FUNCTION_BLOCK StopPointLogic (* Basic Function Block Type *)
  (* Standard: 61499-2 *)
  (* Version 0.0, 11/22/2026, Schneider Electric, First version *)
  PACKAGE Main;
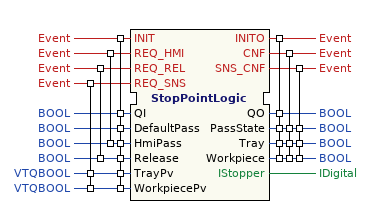
  EVENT_INPUT
    INIT WITH QI, DefaultPass, HmiPass, Release, TrayPv, WorkpiecePv; (* Initialization Request *)
    REQ_HMI WITH HmiPass; (* Update pass-through command from HMI SetBool *)
    REQ_REL WITH Release; (* Update external release request *)
    REQ_SNS WITH TrayPv, WorkpiecePv; (* Update tray and workpiece sensor values *)
  END_EVENT
  EVENT_OUTPUT
    INITO WITH QO, PassState, Tray, Workpiece; (* Initialization Confirm *)
    CNF WITH PassState, Tray, Workpiece; (* Pass-through state confirmation *)
    SNS_CNF WITH Tray, Workpiece, PassState; (* Sensor confirmation *)
  END_EVENT
  VAR_INPUT
    QI : BOOL := TRUE; (* Input event qualifier *)
    DefaultPass : BOOL := FALSE; (* Startup pass-through state (FALSE=Block, TRUE=Pass) *)
    HmiPass : BOOL := FALSE; (* HMI pass-through command *)
    Release : BOOL := FALSE; (* External temporary release input *)
    TrayPv : VTQBOOL; (* Tray-present digital input process value *)
    WorkpiecePv : VTQBOOL; (* Workpiece-present digital input process value *)
  END_VAR
  VAR_OUTPUT
    QO : BOOL; (* Output event qualifier *)
    PassState : BOOL; (* Effective pass-through state (TRUE=stopper down, FALSE=stopper up) *)
    Tray : BOOL; (* Tray present at stop point *)
    Workpiece : BOOL; (* Workpiece present on tray *)
  END_VAR
  PLUGS
    IStopper : IDigital; (* Remote setpoint adapter for Stopper DigitalOutput *)
  END_PLUGS
  VAR
    cmdPass : BOOL := FALSE; (* Latched pass-through command *)
    firstFbDone : BOOL := FALSE; (* Initial REQ_FB sync completed *)
    prevTrack : BOOL := FALSE; (* Previous Track state from Stopper *)
    targetInt : INT := 0; (* Target integer setpoint (0=Block/Up, 1=Pass/Down) *)
  END_VAR
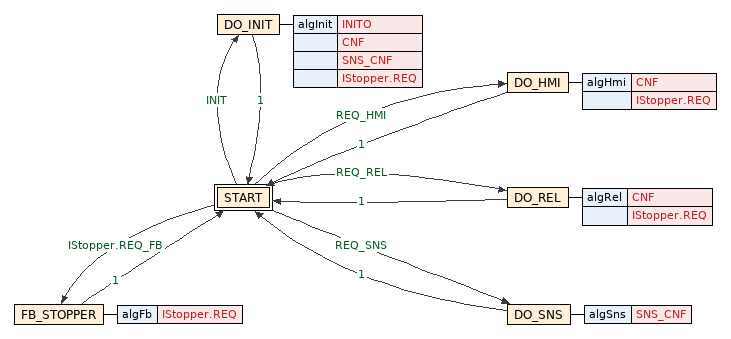
  EC_STATES
    START; (* Initial State *)
    DO_INIT : algInit -> INITO, -> CNF, -> SNS_CNF, -> IStopper.REQ;
    DO_HMI : algHmi -> CNF, -> IStopper.REQ;
    DO_REL : algRel -> CNF, -> IStopper.REQ;
    DO_SNS : algSns -> SNS_CNF;
    FB_STOPPER : algFb -> IStopper.REQ;
  END_STATES
  EC_TRANSITIONS
    START TO DO_INIT := INIT;
    DO_INIT TO START := 1;
    START TO DO_HMI := REQ_HMI;
    DO_HMI TO START := 1;
    START TO DO_REL := REQ_REL;
    DO_REL TO START := 1;
    START TO DO_SNS := REQ_SNS;
    DO_SNS TO START := 1;
    START TO FB_STOPPER := IStopper.REQ_FB;
    FB_STOPPER TO START := 1;
  END_TRANSITIONS
  ALGORITHM algInit IN ST: (* Initialize stop point state from DefaultPass and current sensors *)
QO := QI;
cmdPass := DefaultPass;
PassState := cmdPass OR Release;
IF PassState THEN
	targetInt := 1;
ELSE
	targetInt := 0;
END_IF;

IStopper.Value.value := targetInt;
IStopper.Value.quality := 16#0;

Tray := TrayPv.value;
Workpiece := WorkpiecePv.value;
  END_ALGORITHM
  ALGORITHM algHmi IN ST: (* Update pass-through setpoint from HMI command *)
cmdPass := HmiPass;
PassState := cmdPass OR Release;
IF PassState THEN
	targetInt := 1;
ELSE
	targetInt := 0;
END_IF;

IStopper.Value.value := targetInt;
IStopper.Value.quality := 16#0;
  END_ALGORITHM
  ALGORITHM algRel IN ST: (* Update pass-through setpoint from external release signal *)
PassState := cmdPass OR Release;
IF PassState THEN
	targetInt := 1;
ELSE
	targetInt := 0;
END_IF;

IStopper.Value.value := targetInt;
IStopper.Value.quality := 16#0;
  END_ALGORITHM
  ALGORITHM algSns IN ST: (* Forward VTQBOOL sensor values as clean BOOL outputs *)
Tray := TrayPv.value;
Workpiece := WorkpiecePv.value;
  END_ALGORITHM
  ALGORITHM algFb IN ST: (* Sync Stopper remote setpoint on first feedback or return to Program Remote *)
IStopper.REQ := FALSE;
IF (NOT IStopper.Track) AND ((NOT firstFbDone) OR prevTrack) THEN
	firstFbDone := TRUE;
	PassState := cmdPass OR Release;
	IF PassState THEN
		targetInt := 1;
	ELSE
		targetInt := 0;
	END_IF;
	IStopper.Value.value := targetInt;
	IStopper.Value.quality := 16#0;
	IStopper.REQ := TRUE;
END_IF;
prevTrack := IStopper.Track;
  END_ALGORITHM
END_FUNCTION_BLOCK
